Fanuc KAREL source: kt00728.KL

-- PROVISIONAL review KL for V940-1; original PC SHA256 8fb61bba72d05f73fc90918e50f220668c9cfd514325958beb80e668c186fb76
-- Incomplete behavior may be omitted. Consult companion uncertainty JSON. Do not deploy.
PROGRAM KT00728
%NOLOCKGROUP
VAR
  OUT : BOOLEAN
-- UNRESOLVED_DECL C1 type=00001c
-- UNRESOLVED_DECL C2 type=00001c
BEGIN
  -- V9_ZERO_TABLE_METADATA_HINT layout=0001; no indexed target words; source/name/runtime held
  -- UNRESOLVED_PC offsets 5-15; opcodes 9D,22,A5
  -- UNRESOLVED_PC offsets 20-30; opcodes 9C,22,A5
  -- UNRESOLVED_PC offsets 35-45; opcodes 9D,22,A5
  -- UNRESOLVED_PC offsets 50-60; opcodes 9C,22,A5
  -- UNRESOLVED_PC offsets 65-80; opcodes 22,63,23
  -- UNRESOLVED_PC offsets 85-89; opcodes 7F
END KT00728
